FUNCTION_BLOCK basicGradeamento (* Logica do gradeamento mecanizado (painel Vibropac, Modbus TCP Inovaisa) *)
  (* Standard: 61499-2 *)
  (* Version 1.1, 22/10/2026, Hidryco, Hidryco, 1.1: REQ_GERADOR (geradorHabilita, stsGerador): com a planta nos geradores e a grade nao liberada o ciclo remoto (4001) fica em 0 (stsBloqueioGerador). 1.0: ciclo remoto 4001, reset 4002 (3 s), setpoints 4003/4004 em % (x10 no CLP), leitura 4005..4018, niveis em % *)
  PACKAGE Hidryco.HidrycoLib;
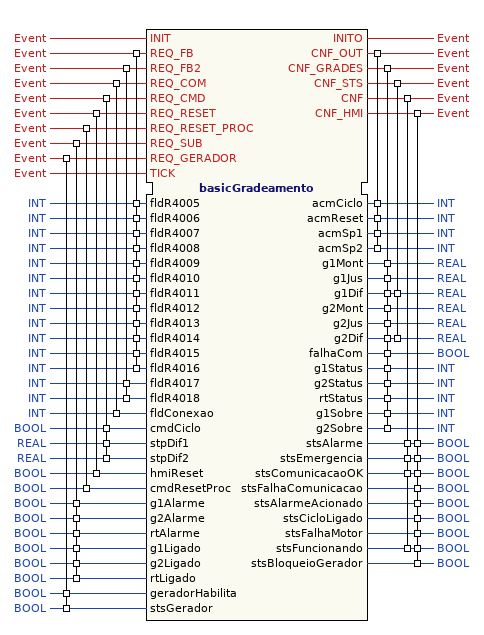
  EVENT_INPUT
    INIT; (* Inicializacao *)
    REQ_FB WITH fldR4005, fldR4006, fldR4007, fldR4008, fldR4009, fldR4010, fldR4011, fldR4012, fldR4013, fldR4014, fldR4015, fldR4016; (* Leitura Modbus 4005..4016 *)
    REQ_FB2 WITH fldR4017, fldR4018; (* Leitura Modbus 4017..4018 *)
    REQ_COM WITH fldConexao; (* Status da conexao Modbus (connStatusInt) *)
    REQ_CMD WITH cmdCiclo, stpDif1, stpDif2; (* Grade_Status1: ciclo remoto e setpoints *)
    REQ_RESET WITH hmiReset; (* IHM: reset (E_RESET_FALHAS_PROCESSO / cmdResetFalhas) *)
    REQ_RESET_PROC WITH cmdResetProc; (* Processo: reset *)
    REQ_SUB WITH g1Alarme, g2Alarme, rtAlarme, g1Ligado, g2Ligado, rtLigado; (* Status das grades e da rosca *)
    REQ_GERADOR WITH geradorHabilita, stsGerador; (* Subestacao: planta nos geradores e liberacao da grade *)
    TICK; (* Base de tempo de 1 s *)
  END_EVENT
  EVENT_OUTPUT
    INITO; (* Inicializacao concluida *)
    CNF_OUT WITH acmCiclo, acmReset, acmSp1, acmSp2; (* Escrita Modbus 4001..4004 *)
    CNF_GRADES WITH g1Mont, g1Jus, g1Dif, g2Mont, g2Jus, g2Dif, falhaCom, g1Status, g2Status, rtStatus, g1Sobre, g2Sobre; (* Leitura para as grades, a rosca e os sensores (na mudanca e a cada 1 s) *)
    CNF_STS WITH g1Dif, g2Dif; (* Diferenciais para o Grade_Status1 (no maximo 1 vez por segundo) *)
    CNF WITH stsAlarme, stsEmergencia, stsComunicacaoOK, stsFuncionando; (* Status para o processo *)
    CNF_HMI WITH stsAlarme, stsEmergencia, stsComunicacaoOK, stsFalhaComunicacao, stsAlarmeAcionado, stsCicloLigado, stsFalhaMotor, stsFuncionando, stsBloqueioGerador; (* Status para a IHM e alarmes *)
  END_EVENT
  VAR_INPUT
    fldR4005 : INT; (* Registro 4005 *)
    fldR4006 : INT; (* Registro 4006 *)
    fldR4007 : INT; (* Registro 4007 *)
    fldR4008 : INT; (* Registro 4008 *)
    fldR4009 : INT; (* Registro 4009 *)
    fldR4010 : INT; (* Registro 4010 *)
    fldR4011 : INT; (* Registro 4011 *)
    fldR4012 : INT; (* Registro 4012 *)
    fldR4013 : INT; (* Registro 4013 *)
    fldR4014 : INT; (* Registro 4014 *)
    fldR4015 : INT; (* Registro 4015 *)
    fldR4016 : INT; (* Registro 4016 *)
    fldR4017 : INT; (* Registro 4017 *)
    fldR4018 : INT; (* Registro 4018 *)
    fldConexao : INT; (* connStatusInt (1 = online) *)
    cmdCiclo : BOOL; (* CMD_LIGA_CICLO_REMOTO *)
    stpDif1 : REAL; (* STP_DIFERENCIAL_NIVEL_GRADE1 (mm) *)
    stpDif2 : REAL; (* STP_DIFERENCIAL_NIVEL_GRADE2 (mm) *)
    hmiReset : BOOL; (* IHM: reset *)
    cmdResetProc : BOOL; (* Processo: reset *)
    g1Alarme : BOOL;
    g2Alarme : BOOL;
    rtAlarme : BOOL;
    g1Ligado : BOOL;
    g2Ligado : BOOL;
    rtLigado : BOOL;
    geradorHabilita : BOOL; (* Grade liberada para operar com a planta nos geradores *)
    stsGerador : BOOL; (* TRUE = planta alimentada pelos geradores *)
  END_VAR
  VAR_OUTPUT
    acmCiclo : INT; (* Registro 4001: 1 liga ciclo remoto, 0 desliga *)
    acmReset : INT; (* Registro 4002: 1 reseta falhas (pulso de 3 s) *)
    acmSp1 : INT; (* Registro 4003: setpoint diferencial grade 1 (0-1000 = 0-100 %) *)
    acmSp2 : INT; (* Registro 4004: setpoint diferencial grade 2 (0-1000 = 0-100 %) *)
    g1Mont : REAL; (* Nivel montante grade 1 LSH1 (%) *)
    g1Jus : REAL; (* Nivel jusante grade 1 LSH2 (%) *)
    g1Dif : REAL; (* Nivel diferencial grade 1 (%) *)
    g2Mont : REAL; (* Nivel montante grade 2 LSH3 (%) *)
    g2Jus : REAL; (* Nivel jusante grade 2 LSH4 (%) *)
    g2Dif : REAL; (* Nivel diferencial grade 2 (%) *)
    falhaCom : BOOL; (* Sem comunicacao com o painel *)
    g1Status : INT; (* Registro 4007 *)
    g2Status : INT; (* Registro 4008 *)
    rtStatus : INT; (* Registro 4009 *)
    g1Sobre : INT; (* Registro 4010 *)
    g2Sobre : INT; (* Registro 4011 *)
    stsAlarme : BOOL; (* Algum alarme do gradeamento (comunicacao, painel, emergencia, motores) *)
    stsEmergencia : BOOL; (* Botao de emergencia do painel acionado (4006) *)
    stsComunicacaoOK : BOOL; (* Comunicacao Modbus com o CLP do painel OK *)
    stsFalhaComunicacao : BOOL; (* Falha de comunicacao com o CLP do painel *)
    stsAlarmeAcionado : BOOL; (* Alarme acionado no painel (4005) *)
    stsCicloLigado : BOOL; (* Comando de ciclo remoto ligado (4001 = 1) *)
    stsFalhaMotor : BOOL; (* Grade ou rosca em falha ou sobretorque *)
    stsFuncionando : BOOL; (* Alguma grade ou a rosca funcionando *)
    stsBloqueioGerador : BOOL; (* Ciclo bloqueado: planta nos geradores e grade nao liberada *)
  END_VAR
  VAR
    initDone : BOOL;
    comRecebido : BOOL;
    fbRecebido : BOOL;
    fb2Recebido : BOOL;
    tReset : INT; (* Segundos restantes do pulso de reset *)
    tEnvio : INT;
    primeiro : BOOL := TRUE;
    oldCiclo : INT := -1;
    oldReset : INT := -1;
    oldSp1 : INT := -1;
    oldSp2 : INT := -1;
    sigG : DINT;
    oldSigG : DINT := -1;
    sig : INT;
    oldSig : INT := -1;
    oldDif1 : REAL := -1.0;
    oldDif2 : REAL := -1.0;
    bBloqGerador : BOOL; (* Planta nos geradores e grade nao liberada *)
  END_VAR
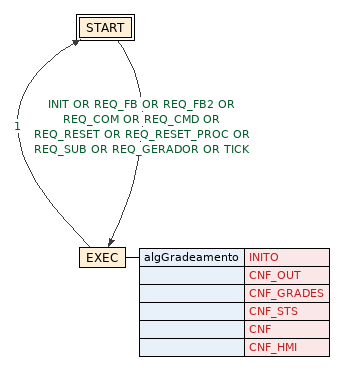
  EC_STATES
    START; (* Estado inicial *)
    EXEC : algGradeamento -> INITO, -> CNF_OUT, -> CNF_GRADES, -> CNF_STS, -> CNF, -> CNF_HMI; (* Executa a logica; o algoritmo decide quais eventos saem *)
  END_STATES
  EC_TRANSITIONS
    START TO EXEC := INIT OR REQ_FB OR REQ_FB2 OR REQ_COM OR REQ_CMD OR REQ_RESET OR REQ_RESET_PROC OR REQ_SUB OR REQ_GERADOR OR TICK;
    EXEC TO START := 1;
  END_TRANSITIONS
  ALGORITHM algGradeamento IN ST: (* Logica completa (um unico algoritmo) *)
(* =====================================================================
   basicGradeamento v1.0 - logica do CAT Gradeamento_Inovaisa (HidrycoLib)
   Painel Vibropac PV-35524 (CLP TM241, tabela Modbus TCP Inovaisa Rev.B):
   4001 liga/desliga ciclo remoto, 4002 reset, 4003/4004 setpoint do
   diferencial de nivel das grades (mm), 4005 alarme,
   4006 emergencia, 4007/4008 grades (0 parado, 1 avante, 2 reverso,
   3 falha), 4009 rosca (0 parado, 1 funcionando, 2 falha), 4010/4011
   sobretorque, 4013..4018 niveis montante/jusante/diferencial (mm).
   O painel tem a propria logica (limpeza pelo diferencial, reverso,
   rosca); o CLP da planta liga/desliga o ciclo, manda os setpoints e le.
   Regras:
   - escrita a cada 5 s e na mudanca (o painel guarda o ultimo valor);
   - reset (IHM ou processo): 4002 = 1 por 3 s;
   - niveis e setpoints de diferencial em mm, sem conversao (valor do registrador = mm);
   - sem comunicacao: estados zerados, sensores em falha de comunicacao.
   ===================================================================== *)
INITO      := FALSE;
CNF_OUT    := FALSE;
CNF_GRADES := FALSE;
CNF_STS    := FALSE;
CNF        := FALSE;
CNF_HMI    := FALSE;
IF REQ_COM THEN
    comRecebido := TRUE;
END_IF;
IF REQ_FB THEN
    fbRecebido := TRUE;
END_IF;
IF REQ_FB2 THEN
    fb2Recebido := TRUE;
END_IF;
IF INIT THEN
    initDone := TRUE;
    INITO := TRUE;
END_IF;
IF NOT initDone THEN
    RETURN;
END_IF;

(* ---- 1. Comunicacao e decodificacao ---- *)
stsComunicacaoOK := comRecebido AND fbRecebido AND fb2Recebido AND (fldConexao = 1);
stsFalhaComunicacao := NOT stsComunicacaoOK;
falhaCom := stsFalhaComunicacao;
IF stsComunicacaoOK THEN
    stsAlarmeAcionado := fldR4005 <> 0;
    stsEmergencia := fldR4006 <> 0;
    g1Status := fldR4007;
    g2Status := fldR4008;
    rtStatus := fldR4009;
    g1Sobre := fldR4010;
    g2Sobre := fldR4011;
    g1Mont := INT_TO_REAL(fldR4013);     (* mm *)
    g1Jus  := INT_TO_REAL(fldR4014);
    g1Dif  := INT_TO_REAL(fldR4015);
    g2Mont := INT_TO_REAL(fldR4016);
    g2Jus  := INT_TO_REAL(fldR4017);
    g2Dif  := INT_TO_REAL(fldR4018);
ELSE
    stsAlarmeAcionado := FALSE;
    stsEmergencia := FALSE;
    g1Status := 0; g2Status := 0; rtStatus := 0; g1Sobre := 0; g2Sobre := 0;
    g1Mont := 0.0; g1Jus := 0.0; g1Dif := 0.0; g2Mont := 0.0; g2Jus := 0.0; g2Dif := 0.0;
END_IF;

(* ---- 2. Comandos (4001..4004) e reset ---- *)
(* planta nos geradores e grade nao liberada na Subestacao: ciclo remoto em 0 *)
bBloqGerador := stsGerador AND NOT geradorHabilita;
stsBloqueioGerador := bBloqGerador;
stsCicloLigado := cmdCiclo AND NOT bBloqGerador;
IF (REQ_RESET AND hmiReset) OR (REQ_RESET_PROC AND cmdResetProc) THEN
    tReset := 3;
END_IF;
IF TICK AND (tReset > 0) THEN
    tReset := tReset - 1;
END_IF;
IF cmdCiclo AND NOT bBloqGerador THEN
    acmCiclo := 1;
ELSE
    acmCiclo := 0;
END_IF;
IF tReset > 0 THEN
    acmReset := 1;
ELSE
    acmReset := 0;
END_IF;
acmSp1 := REAL_TO_INT(LIMIT(0.0, stpDif1, 32767.0));    (* mm *)
acmSp2 := REAL_TO_INT(LIMIT(0.0, stpDif2, 32767.0));
IF TICK THEN
    tEnvio := tEnvio + 1;
END_IF;
IF primeiro OR (acmCiclo <> oldCiclo) OR (acmReset <> oldReset) OR (acmSp1 <> oldSp1) OR (acmSp2 <> oldSp2) OR (tEnvio >= 5) THEN
    CNF_OUT := TRUE;
    tEnvio := 0;
    oldCiclo := acmCiclo; oldReset := acmReset; oldSp1 := acmSp1; oldSp2 := acmSp2;
END_IF;

(* ---- 3. Para as grades, a rosca e os sensores: na mudanca do estado e a cada 1 s (niveis) ---- *)
sigG := INT_TO_DINT(g1Status) + INT_TO_DINT(g2Status) * 8 + INT_TO_DINT(rtStatus) * 64 + INT_TO_DINT(g1Sobre) * 512 + INT_TO_DINT(g2Sobre) * 1024;
IF falhaCom THEN sigG := sigG + 4096; END_IF;
IF primeiro OR TICK OR (sigG <> oldSigG) THEN
    CNF_GRADES := TRUE;
END_IF;
oldSigG := sigG;
IF TICK AND ((g1Dif <> oldDif1) OR (g2Dif <> oldDif2)) THEN
    CNF_STS := TRUE;
    oldDif1 := g1Dif; oldDif2 := g2Dif;
END_IF;

(* ---- 4. Alarme geral ---- *)
stsFalhaMotor := g1Alarme OR g2Alarme OR rtAlarme;
stsFuncionando := g1Ligado OR g2Ligado OR rtLigado;
stsAlarme := stsFalhaComunicacao OR stsAlarmeAcionado OR stsEmergencia OR stsFalhaMotor;

(* ---- 5. Eventos ---- *)
sig := 0;
IF stsComunicacaoOK THEN sig := sig + 1; END_IF;
IF stsAlarmeAcionado THEN sig := sig + 2; END_IF;
IF stsEmergencia THEN sig := sig + 4; END_IF;
IF stsCicloLigado THEN sig := sig + 8; END_IF;
IF stsFalhaMotor THEN sig := sig + 16; END_IF;
IF stsFuncionando THEN sig := sig + 32; END_IF;
IF stsAlarme THEN sig := sig + 64; END_IF;
IF stsBloqueioGerador THEN sig := sig + 128; END_IF;
IF primeiro OR REQ_RESET OR (sig <> oldSig) THEN
    CNF_HMI := TRUE;
    CNF := TRUE;
END_IF;
oldSig := sig;
primeiro := FALSE;
  END_ALGORITHM
END_FUNCTION_BLOCK
